(* CODESYS project Example11_PLC.project

Project tree, tasks and I/O mapping:
  Device : CODESYS Control Win V3, 3S - Smart Software Solutions GmbH, order no. 305021, version 3.5.7.0
    application Application
      libraries: Standard, * (System)
      task MainTask (cyclic, interval t#20ms, priority 1) calls PLC_PRG
      program PLC_PRG [ST]
      global variables GVL
      function block FB_G4LTL [ST]
    Ethernet : Ethernet, 3S - Smart Software Solutions GmbH, version 3.5.7.0
      Modbus_TCP_Master : Modbus TCP Master, 3S - Smart Software Solutions GmbH, version 3.5.6.0
          settings: AutoReconnect = TRUE
        Modbus_TCP_Slave : Modbus TCP Slave, 3S - Smart Software Solutions GmbH, version 3.5.7.0
            settings: Unit-ID = 1; IPAddress = [127, 0, 0, 1]; Channel 0.Function Code = 4; Channel 0.Read Offset = 16#0000; Channel 0.Read Length = 1; Channel 0.Write Offset = 0; Channel 0.Write Length = 0; Channel 0.Cycle Time = 100; Channel 1.Function Code = 4; Channel 1.Read Offset = 16#0001; Channel 1.Read Length = 1; Channel 1.Write Offset = 0; Channel 1.Write Length = 0; Channel 1.Cycle Time = 100; Channel 2.Function Code = 4; Channel 2.Read Offset = 16#0002; Channel 2.Read Length = 1; Channel 2.Write Offset = 0; Channel 2.Write Length = 0; Channel 2.Cycle Time = 100; Channel 3.Function Code = 4; Channel 3.Read Offset = 16#0003; Channel 3.Read Length = 1; Channel 3.Write Offset = 0; Channel 3.Write Length = 0; Channel 3.Cycle Time = 100; Channel 4.Function Code = 4; Channel 4.Read Offset = 16#0004; Channel 4.Read Length = 1; Channel 4.Write Offset = 0; Channel 4.Write Length = 0; Channel 4.Cycle Time = 100; Channel 5.Function Code = 6; Channel 5.Read Offset = 0; Channel 5.Read Length = 0; Channel 5.Write Offset = 16#0000; Channel 5.Write Length = 1; Channel 5.Cycle Time = 100; Channel 6.Function Code = 6; Channel 6.Read Offset = 0;
              Channel 6.Read Length = 0; Channel 6.Write Offset = 16#0002; Channel 6.Write Length = 1; Channel 6.Cycle Time = 100; Channel 7.Function Code = 6; Channel 7.Read Offset = 0; Channel 7.Read Length = 0; Channel 7.Write Offset = 16#0003; Channel 7.Write Length = 1; Channel 7.Cycle Time = 100; Channel 8.Function Code = 6; Channel 8.Read Offset = 0; Channel 8.Read Length = 0; Channel 8.Write Offset = 16#0004; Channel 8.Write Length = 1; Channel 8.Cycle Time = 100; Channel 9.Function Code = 6; Channel 9.Read Offset = 0; Channel 9.Read Length = 0; Channel 9.Write Offset = 16#0001; Channel 9.Write Length = 1; Channel 9.Cycle Time = 100; Channel 10.Function Code = 4; Channel 10.Read Offset = 16#0005; Channel 10.Read Length = 1; Channel 10.Write Offset = 0; Channel 10.Write Length = 0; Channel 10.Cycle Time = 100
            input  Application.dIn0 : BOOL  // Channel 0.Channel 0.Bit0
            input  Application.dIn1 : BOOL  // Channel 1.Channel 1.Bit0
            input  Application.dIn2 : BOOL  // Channel 2.Channel 2.Bit0
            input  Application.dIn3 : BOOL  // Channel 3.Channel 3.Bit0
            input  Application.dIn4 : BOOL  // Channel 4.Channel 4.Bit0
            output Application.dOut0 : BOOL  // Channel 5.Channel 5.Bit0
            output Application.dOut2 : BOOL  // Channel 6.Channel 6.Bit0
            output Application.dOut3 : BOOL  // Channel 7.Channel 7.Bit0
            output Application.dOut4 : BOOL  // Channel 8.Channel 8.Bit0
            output Application.dOut1 : BOOL  // Channel 9.Channel 9.Bit0
            input  Application.dIn5 : BOOL  // Channel 10.Channel 10.Bit0
            unmapped channels: Channel 0, Channel 1, Channel 2, Channel 3, Channel 4, Channel 5, Channel 6, Channel 7, Channel 8, Channel 9, Channel 10
*)

// Device/Application/GVL
VAR_GLOBAL
	
dIn0 : BOOL;
dIn1 : BOOL;
dIn2 : BOOL;
dIn3 : BOOL;
dIn4 : BOOL;
dIn5 : BOOL;

dOut0 : BOOL;
dOut1 : BOOL; 
dOut2 : BOOL; 
dOut3 : BOOL; 
dOut4 : BOOL; 
END_VAR

// Device/Application/PLC_PRG
PROGRAM PLC_PRG

VAR 
	fb: FB_G4LTL;
END_VAR


// Direct looping
// Assign pins (from global variable to function block) 
fb.x1 := dIn0;
fb.x2 := dIn1;

// Assign pins (from function block to global variable)
dOut0 := fb.y0;
dOut1 := fb.y1;
dOut2 := fb.y2;

// Run the function block
fb();

END_PROGRAM

// Device/Application/FB_G4LTL
FUNCTION_BLOCK FB_G4LTL

   (* Variable definition *)
   VAR_INPUT
      x1	: BOOL;
      x2	: BOOL;
   END_VAR
   VAR_OUTPUT
      y0	: BOOL;
      y1	: BOOL;
      y2	: BOOL;
   END_VAR
   VAR
   (* The total number of states equals to 3 *)
      cstate42	: LINT := 0;
   END_VAR

 (* Control logic *)
CASE cstate42 OF
0:
    IF ((x1 = TRUE) AND  (x2 = FALSE)) THEN 
        cstate42 := 12; y0 := TRUE; y1 := TRUE; y2 := FALSE;  
    ELSIF ((x1 = FALSE) AND  ( TRUE )) THEN 
        cstate42 := 7; y0 := FALSE; y1 := FALSE; y2 := TRUE;  
    ELSIF ((x1 = TRUE) AND  (x2 = TRUE)) THEN 
        cstate42 := 14; y0 := FALSE; y1 := TRUE; y2 := FALSE;  
    END_IF;
7:
    IF ((x1 = TRUE) AND  (x2 = FALSE)) THEN 
        cstate42 := 12; y0 := TRUE; y1 := TRUE; y2 := FALSE;  
    ELSIF ((x1 = FALSE) AND  ( TRUE )) THEN 
        cstate42 := 7; y0 := FALSE; y1 := FALSE; y2 := TRUE;  
    ELSIF ((x1 = TRUE) AND  (x2 = TRUE)) THEN 
        cstate42 := 14; y0 := FALSE; y1 := TRUE; y2 := FALSE;  
    END_IF;
14:
    IF ((x1 = TRUE) AND  (x2 = FALSE)) THEN 
        cstate42 := 12; y0 := TRUE; y1 := TRUE; y2 := FALSE;  
    ELSIF ((x1 = FALSE) AND  (x2 = FALSE)) OR ((x1 = TRUE) AND  (x2 = TRUE)) THEN 
        cstate42 := 14; y0 := FALSE; y1 := TRUE; y2 := FALSE;  
    ELSIF ((x1 = FALSE) AND  (x2 = TRUE)) THEN 
        cstate42 := 7; y0 := FALSE; y1 := FALSE; y2 := TRUE;  
    END_IF;
12:
    IF (( TRUE ) AND  (x2 = FALSE)) THEN 
        cstate42 := 12; y0 := TRUE; y1 := TRUE; y2 := FALSE;  
    ELSIF ((x1 = FALSE) AND  (x2 = TRUE)) THEN 
        cstate42 := 7; y0 := FALSE; y1 := FALSE; y2 := TRUE;  
    ELSIF ((x1 = TRUE) AND  (x2 = TRUE)) THEN 
        cstate42 := 14; y0 := FALSE; y1 := TRUE; y2 := FALSE;  
    END_IF;
END_CASE;

END_FUNCTION_BLOCK
